Fanuc KAREL source: kd00052.KL

PROGRAM KD00052
%STACKSIZE=65535
%PRIORITY=65535
%NOLOCKGROUP
VAR
I : INTEGER
J : INTEGER
B : BOOLEAN
R : REAL
S : STRING[80]
P : POSITION
BEGIN
-- UNRESOLVED_PC line 12 opcodes [01 22 1C 06 82 03 9D 2E 51 9D 12 9D 1B 9D 13 04 0B] marker_code=0
END KD00052
